Fanuc KAREL source: kt00533.KL

-- PROVISIONAL review KL for V940-1; original PC SHA256 153658f47573de89d63464450a6328024e6033c27bd5afd4d9bb793dcf41e569
-- Incomplete behavior may be omitted. Consult companion uncertainty JSON. Do not deploy.
PROGRAM KT00533
%NOLOCKGROUP
VAR
  OUT : BOOLEAN
-- UNRESOLVED_DECL P1 type=000199
-- UNRESOLVED_DECL P2 type=000101
BEGIN
  -- V9_ZERO_TABLE_METADATA_HINT layout=0001; no indexed target words; source/name/runtime held
  -- UNRESOLVED_PC offsets 5-33; opcodes 49,7E,49,AC,23
  -- UNRESOLVED_PC offsets 38-42; opcodes 7F
END KT00533
